(* IEC 61131-3 sources: ISA-88-Bioreactor-Automation-Template-DE-IE/ISA-88-Bioreactor-Automation-Template-DE-IE.fbsdev/TankCycler.iecapp^, 7 files *)

(* ---- CycleComplete.fb.st ---- *)
FUNCTION_BLOCK CycleComplete_FB_ST
VAR_INPUT
    Cycle_Active       : BOOL;
    Fill_Complete      : BOOL;
    Mix_Complete       : BOOL;
    Heat_Complete      : BOOL;
    Discharge_Complete : BOOL;
END_VAR

VAR_OUTPUT
    T1_Cycle_Complete  : BOOL := FALSE;
    Cycle_Reset        : BOOL := FALSE;
END_VAR

// Body logic
IF Cycle_Active AND Fill_Complete AND Mix_Complete AND Heat_Complete AND Discharge_Complete THEN
    T1_Cycle_Complete := TRUE;
    Cycle_Reset := TRUE;   // signal to reset latch in TankCycle_FB
ELSE
    T1_Cycle_Complete := FALSE;
    Cycle_Reset := FALSE;
END_IF;

IF Cycle_Active AND Discharge_Complete THEN
    T1_Cycle_Complete := TRUE;
    Cycle_Active := FALSE;   // reset latch
END_IF;

END_FUNCTION_BLOCK

(* ---- DischargeStage.fb.st ---- *)
FUNCTION_BLOCK DischargeStage_FB_ST
VAR_INPUT
  Cycle_Active     : BOOL;
  Heat_Complete    : BOOL;
END_VAR

VAR_OUTPUT
  T1_Valve_Outlet  : BOOL;
  Discharge_Complete : BOOL;
END_VAR

// implementation here...

IF Cycle_Active AND Heat_Complete THEN
    T1_Valve_Outlet := TRUE;
ELSE
    T1_Valve_Outlet := FALSE;
END_IF;

IF Cycle_Active AND Heat_Complete THEN
    Discharge_Complete := TRUE;
END_IF;

END_FUNCTION_BLOCK

(* ---- FillStage.fb.st ---- *)
FUNCTION_BLOCK FillStage_FB_ST

VAR_INPUT
  Cycle_Active   : BOOL;
  T1_Level_High  : BOOL;
END_VAR

VAR_OUTPUT
  T1_Valve_Inlet : BOOL;
  Fill_Complete  : BOOL;
END_VAR

VAR
END_VAR

// implementation here...
// Fill logic
IF Start_Fill THEN
    Valve_Inlet := NOT Tn_Level_High;
    IF Tn_Level_High THEN
        Fill_Complete := TRUE;
        Valve_Inlet := FALSE;
    END_IF;
ELSE
    Valve_Inlet := FALSE;
    Fill_Complete := FALSE;
END_IF;

END_FUNCTION_BLOCK

(* ---- HeatStage.fb.st ---- *)
FUNCTION_BLOCK HeatStage_FB
VAR_INPUT
  Cycle_Active    : BOOL;
  T1_Mix_Complete : BOOL;
  T1_Temp_Sensor  : INT;
  T1_Temp_Setpoint: INT;
END_VAR

VAR_OUTPUT
  T1_Heater       : BOOL;
  T1_Temp_Alarm   : BOOL;
  Heat_Complete   : BOOL;
END_VAR

// implementation here...

IF Cycle_Active AND T1_Mix_Complete AND (T1_Temp_Sensor < T1_Temp_Setpoint) THEN
    T1_Heater := TRUE;
ELSE
    T1_Heater := FALSE;
END_IF;

IF Cycle_Active AND T1_Mix_Complete AND (T1_Temp_Sensor > T1_Temp_Setpoint) THEN
    T1_Temp_Alarm := TRUE;
ELSE
    T1_Temp_Alarm := FALSE;
END_IF;

IF Cycle_Active AND T1_Mix_Complete AND (T1_Temp_Sensor >= T1_Temp_Setpoint) THEN
    Heat_Complete := TRUE;
END_IF;

END_FUNCTION_BLOCK

(* ---- MixStage.fb.st ---- *)
FUNCTION_BLOCK MixStage_FB
VAR_INPUT
    Cycle_Active  : BOOL;   // latch from TankCycle
    Fill_Complete : BOOL;   // signal from FillStage
END_VAR

VAR_OUTPUT
    Mix_Complete  : BOOL := FALSE; // goes high when mixing done
END_VAR

VAR
END_VAR

IF Cycle_Active AND Fill_Complete THEN
    Mix_Complete := TRUE;
ELSE
    Mix_Complete := FALSE;
END_IF;
// implementation here...

END_FUNCTION_BLOCK

(* ---- TankCycle.fb.st ---- *)
FUNCTION_BLOCK TankCycle_FB_ST
FUNCTION_BLOCK TankCycle_FB_ST
VAR_INPUT
    Start_Cycle       : BOOL;   // trigger to start cycle
    Tn_Level_High     : BOOL;   // tank full sensor
    Tn_Level_Low      : BOOL;   // tank empty sensor
    Tn_Temp_Value     : REAL;   // current temperature
    Tn_Temp_Setpoint  : REAL;   // desired temperature
END_VAR

VAR_OUTPUT
    Valve_Inlet       : BOOL := FALSE;
    Mixer_Motor       : BOOL := FALSE;
    Heater            : BOOL := FALSE;
    Valve_Outlet      : BOOL := FALSE;
    Cycle_Complete    : BOOL := FALSE;
END_VAR
VAR
    Fill_Complete     : BOOL := FALSE;
    Mix_Complete      : BOOL := FALSE;
    Heat_Complete     : BOOL := FALSE;
    Discharge_Complete: BOOL := FALSE;
END_VAR

// implementation here...

// Sequence logic
IF Start_Cycle AND NOT Fill_Complete THEN
    Valve_Inlet := NOT Tn_Level_High;
    IF Tn_Level_High THEN
        Fill_Complete := TRUE;
        Valve_Inlet := FALSE;
    END_IF;
END_IF;

IF Fill_Complete AND NOT Mix_Complete THEN
    Mixer_Motor := TRUE;
    // Example: mixing runs for 10s
    // (replace with TON timer instance in real project)
    Mix_Complete := TRUE; // stub: set after timer
    Mixer_Motor := FALSE;
END_IF;

IF Mix_Complete AND NOT Heat_Complete THEN
    Heater := (Tn_Temp_Value < Tn_Temp_Setpoint);
    IF Tn_Temp_Value >= Tn_Temp_Setpoint THEN
        Heat_Complete := TRUE;
        Heater := FALSE;
    END_IF;
END_IF;

IF Heat_Complete AND NOT Discharge_Complete THEN
    Valve_Outlet := NOT Tn_Level_Low;
    IF Tn_Level_Low THEN
        Discharge_Complete := TRUE;
        Valve_Outlet := FALSE;
    END_IF;
END_IF;

IF Discharge_Complete THEN
    Cycle_Complete := TRUE;
END_IF;

END_FUNCTION_BLOCK

(* ---- PLC_PRG.prg.st ---- *)
PROGRAM PLC_PRG
VAR
    FillStage      : FillStage_FB_ST;
    MixStage       : MixStage_FB_ST;
    HeatStage      : HeatStage_FB_ST;
    DischargeStage : DischargeStage_FB_ST;
    CycleComplete  : CycleComplete_FB_ST;
END_VAR

// implementation here...
// TankCycle orchestrates the sequence
TankCycle(
    Start_Cycle     := GV_TankFarm.Start_Cycle,
    T1_Level_High   := GV_TankFarm.T1_Level_High,
    T1_Level_Low    := GV_TankFarm.T1_Level_Low,
    T1_Temp_Value   := GV_TankFarm.T1_Temp_Sensor,
    T1_Temp_Setpoint:= GV_TankFarm.T1_Temp_Setpoint
);

// FillStage
FillStage(
    Start_Fill    := TankCycle.Cycle_Active,
    Tn_Level_High := GV_TankFarm.T1_Level_High
);

// MixStage
MixStage(
    Cycle_Active  := TankCycle.Cycle_Active,
    Fill_Complete := FillStage.Fill_Complete
);

// HeatStage
HeatStage(
    Cycle_Active     := TankCycle.Cycle_Active,
    Mix_Complete     := MixStage.Mix_Complete,
    Tn_Temp_Value    := GV_TankFarm.T1_Temp_Sensor,
    Tn_Temp_Setpoint := TankCycle.Tn_Temp_Setpoint
);

// DischargeStage
DischargeStage(
    Cycle_Active   := TankCycle.Cycle_Active,
    Heat_Complete  := HeatStage.Heat_Complete,
    Tn_Level_Low   := GV_TankFarm.T1_Level_Low
);

// CycleComplete
CycleComplete(
    Cycle_Active       := TankCycle.Cycle_Active,
    Fill_Complete      := FillStage.Fill_Complete,
    Mix_Complete       := MixStage.Mix_Complete,
    Heat_Complete      := HeatStage.Heat_Complete,
    Discharge_Complete := DischargeStage.Discharge_Complete
);

// Reset logic
IF CycleComplete.Cycle_Reset THEN
    TankCycle.Cycle_Active := FALSE;
END_IF;

END_PROGRAM
